(* IEC 61131-3 sources: plcassist-cli/packages/volt-lsp-iec/test-corpus/bakon-nano/Device/Plc Logic/Application/Library Manager/L_PLCLoggingAccess, 10 files *)

(* ---- GETBOOLEANPROPERTY.fun ---- *)
FUNCTION GETBOOLEANPROPERTY : BOOL
VAR_INPUT
	STKEY : WSTRING;
END_VAR
END_FUNCTION

(* ---- GETCOMPANY.fun ---- *)
FUNCTION GETCOMPANY : WSTRING
END_FUNCTION

(* ---- GETNUMBERPROPERTY.fun ---- *)
FUNCTION GETNUMBERPROPERTY : DINT
VAR_INPUT
	STKEY : WSTRING;
END_VAR
END_FUNCTION

(* ---- GETTEXTPROPERTY.fun ---- *)
FUNCTION GETTEXTPROPERTY : WSTRING
VAR_INPUT
	STKEY : WSTRING;
END_VAR
END_FUNCTION

(* ---- GETTEXTPROPERTY2.fun ---- *)
FUNCTION GETTEXTPROPERTY2 : POINTER TO WSTRING
VAR_INPUT
	STKEY : WSTRING;
END_VAR
END_FUNCTION

(* ---- GETTITLE.fun ---- *)
FUNCTION GETTITLE : WSTRING
END_FUNCTION

(* ---- GETVERSION.fun ---- *)
FUNCTION GETVERSION : VERSION
END_FUNCTION

(* ---- GETVERSIONPROPERTY.fun ---- *)
FUNCTION GETVERSIONPROPERTY : VERSION
VAR_INPUT
	STKEY : WSTRING;
END_VAR
END_FUNCTION

(* ---- L_ADDLOG.fun ---- *)
FUNCTION L_ADDLOG : BOOL
VAR_INPUT
	ESEVERITY : L_TSeverity;
	EFACILITY : L_TFacility;
	SLOGPAYLOAD : STRING(80);
END_VAR
END_FUNCTION

(* ---- L_ADDLOG2.fun ---- *)
FUNCTION L_ADDLOG2 : BOOL
VAR_INPUT
	ESEVERITY : L_TSeverity;
	UDICOMPONENDID : UDINT;
	SLOGPAYLOAD : STRING(80);
	DWERRORID : DWORD;
	STRLANGUAGETABLE : STRING(80);
END_VAR
END_FUNCTION
